// Mitsubishi GX Works2 project: 공개2번(FX)   PLC: FX3U/FX3UC

PROGRAM MAIN
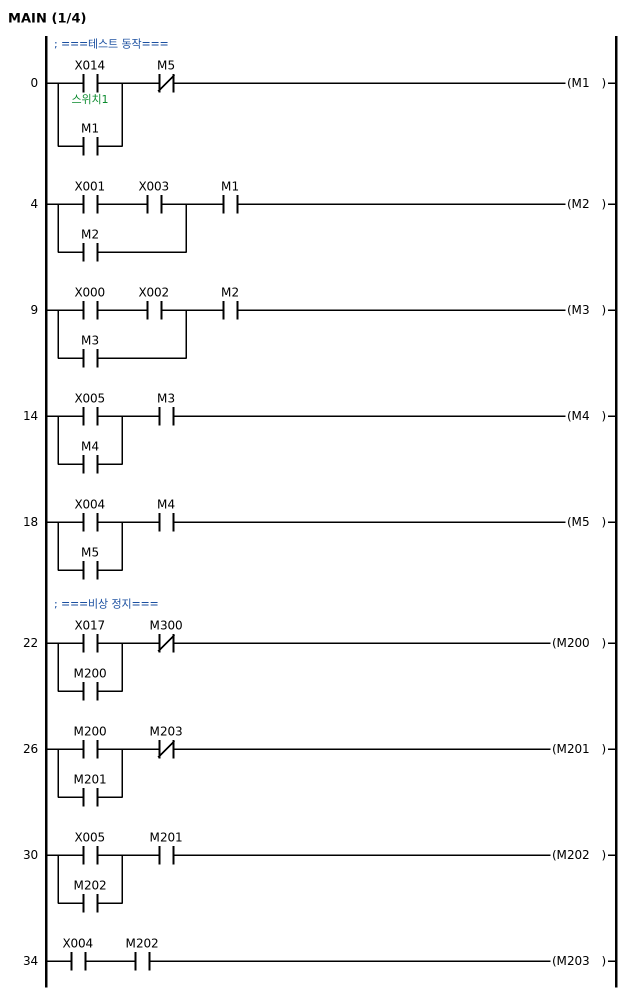
; ===테스트 동작===
0     LD      X014  ; 스위치1
      OR      M1
      ANI     M5
      OUT     M1
4     LD      X001
      AND     X003
      OR      M2
      AND     M1
      OUT     M2
9     LD      X000
      AND     X002
      OR      M3
      AND     M2
      OUT     M3
14    LD      X005
      OR      M4
      AND     M3
      OUT     M4
18    LD      X004
      OR      M5
      AND     M4
      OUT     M5
; ===비상 정지===
22    LD      X017
      OR      M200
      ANI     M300
      OUT     M200
26    LD      M200
      OR      M201
      ANI     M203
      OUT     M201
30    LD      X005
      OR      M202
      AND     M201
      OUT     M202
34    LD      X004
      AND     M202
      OUT     M203
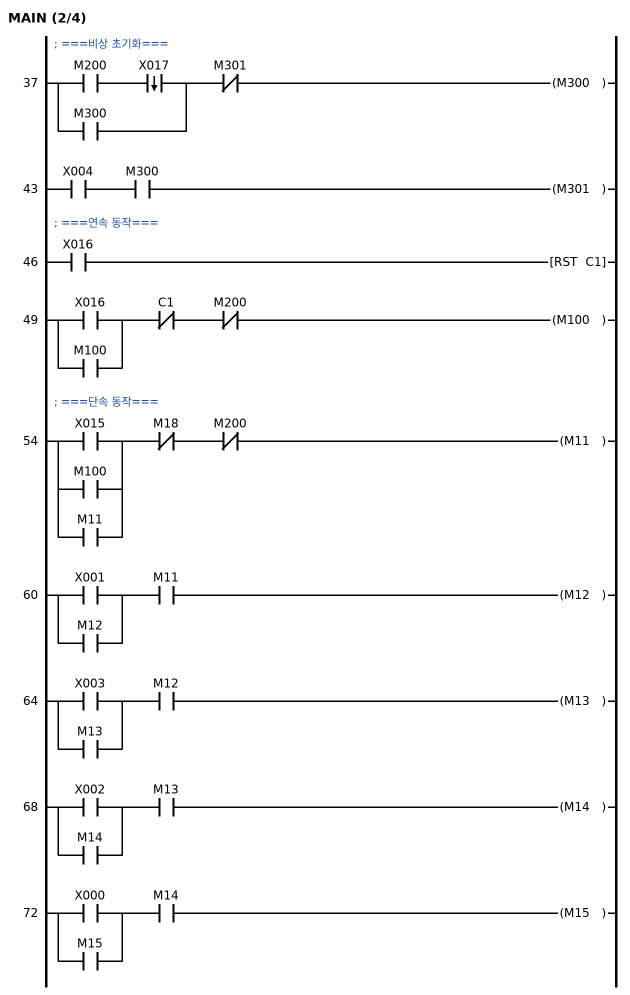
; ===비상 초기화===
37    LD      M200
      ANDF    X017
      OR      M300
      ANI     M301
      OUT     M300
43    LD      X004
      AND     M300
      OUT     M301
; ===연속 동작===
46    LD      X016
      RST     C1
49    LD      X016
      OR      M100
      ANI     C1
      ANI     M200
      OUT     M100
; ===단속 동작===
54    LD      X015
      OR      M100
      OR      M11
      ANI     M18
      ANI     M200
      OUT     M11
60    LD      X001
      OR      M12
      AND     M11
      OUT     M12
64    LD      X003
      OR      M13
      AND     M12
      OUT     M13
68    LD      X002
      OR      M14
      AND     M13
      OUT     M14
72    LD      X000
      OR      M15
      AND     M14
      OUT     M15
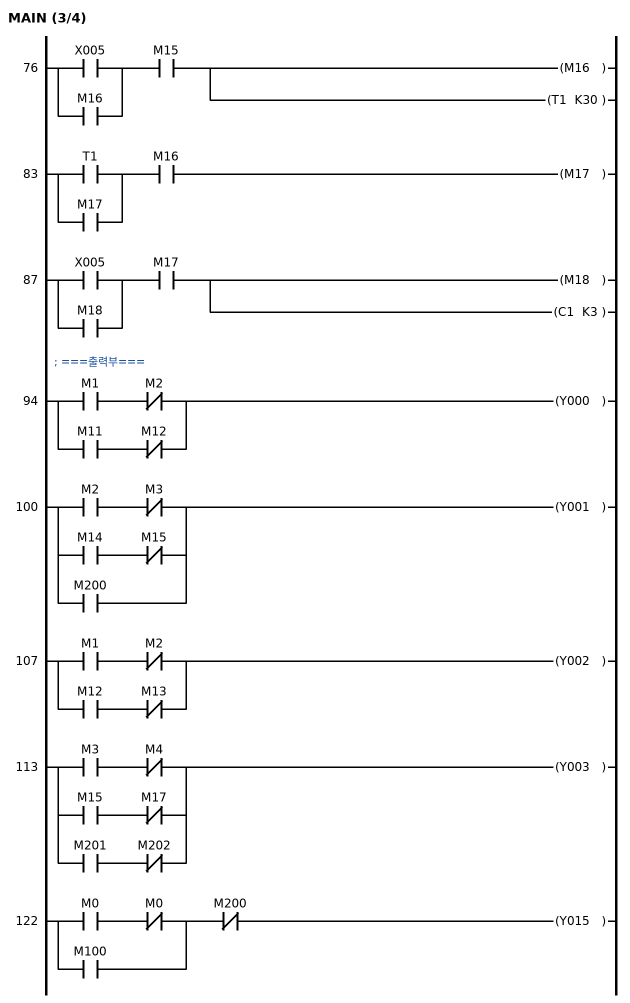
76    LD      X005
      OR      M16
      AND     M15
      OUT     M16
      OUT     T1 K30
83    LD      T1
      OR      M17
      AND     M16
      OUT     M17
87    LD      X005
      OR      M18
      AND     M17
      OUT     M18
      OUT     C1 K3
; ===출력부===
94    LD      M1
      ANI     M2
      LD      M11
      ANI     M12
      ORB
      OUT     Y000
100   LD      M2
      ANI     M3
      LD      M14
      ANI     M15
      ORB
      OR      M200
      OUT     Y001
107   LD      M1
      ANI     M2
      LD      M12
      ANI     M13
      ORB
      OUT     Y002
113   LD      M3
      ANI     M4
      LD      M15
      ANI     M17
      ORB
      LD      M201
      ANI     M202
      ORB
      OUT     Y003
122   LD      M0
      ANI     M0
      OR      M100
      ANI     M200
      OUT     Y015
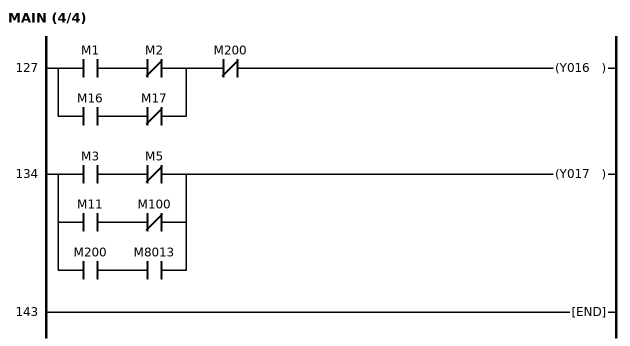
127   LD      M1
      ANI     M2
      LD      M16
      ANI     M17
      ORB
      ANI     M200
      OUT     Y016
134   LD      M3
      ANI     M5
      LD      M11
      ANI     M100
      ORB
      LD      M200
      AND     M8013
      ORB
      OUT     Y017
143   END
END_PROGRAM
